FUNCTION_BLOCK F (* Negative C3: a real lowered TON body, whose state variable a guard reads as a position, so the exemption is lost *)
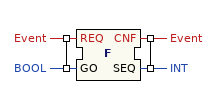
  EVENT_INPUT
    REQ WITH GO;
  END_EVENT
  EVENT_OUTPUT
    CNF WITH SEQ;
  END_EVENT
  VAR_INPUT
    GO : BOOL;
  END_VAR
  VAR_OUTPUT
    SEQ : INT;
  END_VAR
  VAR
    T_STATE : INT;
    T_PREV_IN : BOOL;
    T_Q : BOOL;
    T_START_TIME : TIME;
    NOW : TIME;
  END_VAR
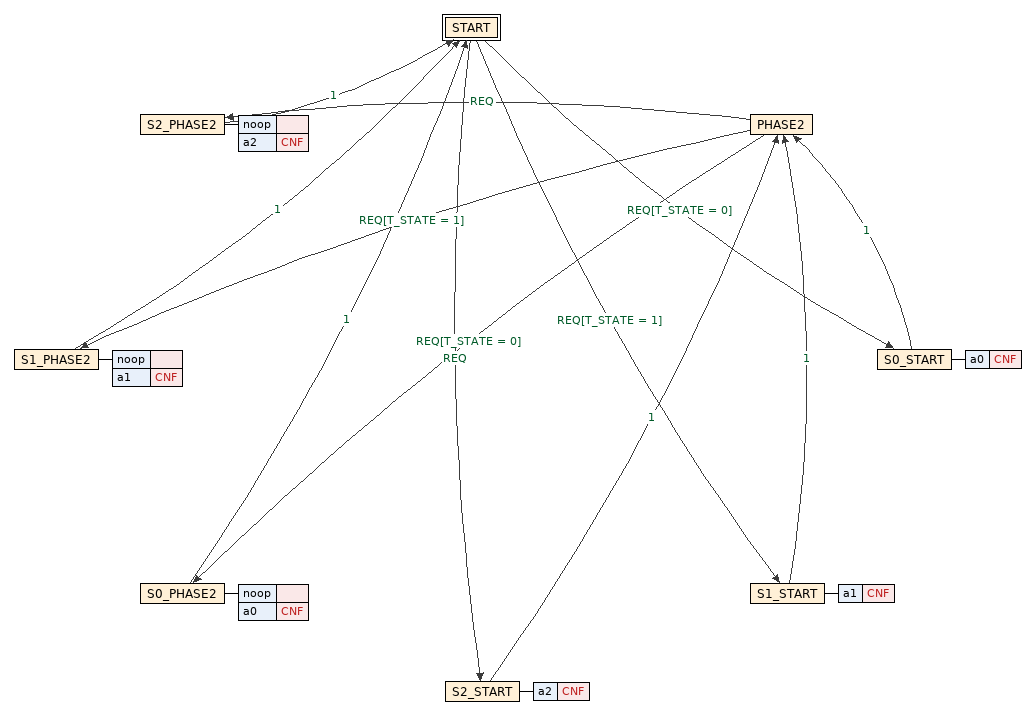
  EC_STATES
    START;
    PHASE2;
    S0_START : a0 -> CNF;
    S1_START : a1 -> CNF;
    S2_START : a2 -> CNF;
    S0_PHASE2 : noop, a0 -> CNF;
    S1_PHASE2 : noop, a1 -> CNF;
    S2_PHASE2 : noop, a2 -> CNF;
  END_STATES
  EC_TRANSITIONS
    START TO S0_START := REQ[T_STATE = 0];
    START TO S1_START := REQ[T_STATE = 1];
    START TO S2_START := REQ;
    PHASE2 TO S0_PHASE2 := REQ[T_STATE = 0];
    PHASE2 TO S1_PHASE2 := REQ[T_STATE = 1];
    PHASE2 TO S2_PHASE2 := REQ;
    S0_START TO PHASE2 := 1;
    S1_START TO PHASE2 := 1;
    S2_START TO PHASE2 := 1;
    S0_PHASE2 TO START := 1;
    S1_PHASE2 TO START := 1;
    S2_PHASE2 TO START := 1;
  END_TRANSITIONS
  ALGORITHM a0 IN ST:
NOW := NOW + T#10ms;
IF (T_STATE = 0) AND NOT T_PREV_IN AND GO THEN
  T_STATE := 1;
  T_START_TIME := NOW;
ELSIF NOT GO THEN
  T_STATE := 0;
ELSIF T_STATE = 1 THEN
  IF T_START_TIME + T#50ms <= NOW THEN
    T_STATE := 2;
    T_Q := TRUE;
  END_IF;
END_IF;
T_PREV_IN := GO;
SEQ := 1;
  END_ALGORITHM
  ALGORITHM a1 IN ST:
SEQ := 2;
  END_ALGORITHM
  ALGORITHM a2 IN ST:
SEQ := 0;
  END_ALGORITHM
  ALGORITHM noop IN ST:
SEQ := SEQ;
  END_ALGORITHM
END_FUNCTION_BLOCK
